Fanuc KAREL source: kb00178.KL

-- PROVISIONAL review KL for V940-1; original PC SHA256 06f796e9ce49e1f32573ac75940a658881bf73b95ad923b0bb311931601ce048
-- Incomplete behavior may be omitted. Consult companion uncertainty JSON. Do not deploy.
PROGRAM KB00178
%NOLOCKGROUP
BEGIN
  -- V9_ZERO_TABLE_METADATA_HINT layout=0002_ascii; no indexed target words; source/name/runtime held
  -- UNRESOLVED_PC offsets 5-12; opcodes 9D,23
  -- UNRESOLVED_PC offsets 17-28; opcodes 2E,23
  -- UNRESOLVED_PC offsets 33-40; opcodes 9D,23
  -- UNRESOLVED_PC offsets 45-67; opcodes 27,22,22,22,31
  -- UNRESOLVED_PC offsets 72-76; opcodes 7F
END KB00178
